// Mitsubishi GX Works2 project: V3 (working)   PLC: FX3U/FX3UC

PROGRAM MAIN
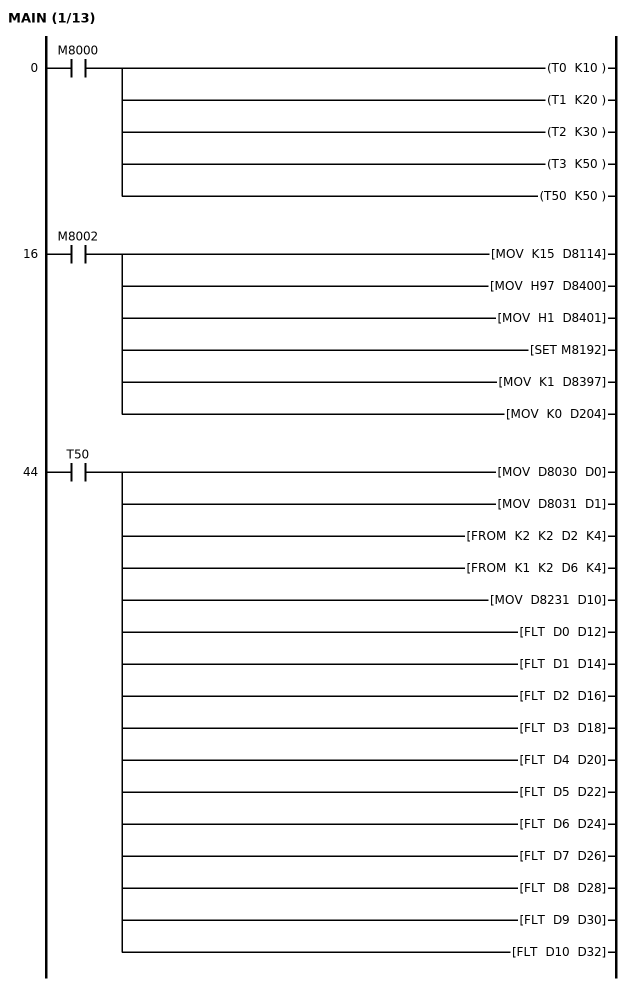
0     LD      M8000
      OUT     T0 K10
      OUT     T1 K20
      OUT     T2 K30
      OUT     T3 K50
      OUT     T50 K50
16    LD      M8002
      MOV     K15 D8114
      MOV     H97 D8400
      MOV     H1 D8401
      SET     M8192
      MOV     K1 D8397
      MOV     K0 D204
44    LD      T50
      MOV     D8030 D0
      MOV     D8031 D1
      FROM    K2 K2 D2 K4
      FROM    K1 K2 D6 K4
      MOV     D8231 D10
      FLT     D0 D12
      FLT     D1 D14
      FLT     D2 D16
      FLT     D3 D18
      FLT     D4 D20
      FLT     D5 D22
      FLT     D6 D24
      FLT     D7 D26
      FLT     D8 D28
      FLT     D9 D30
      FLT     D10 D32
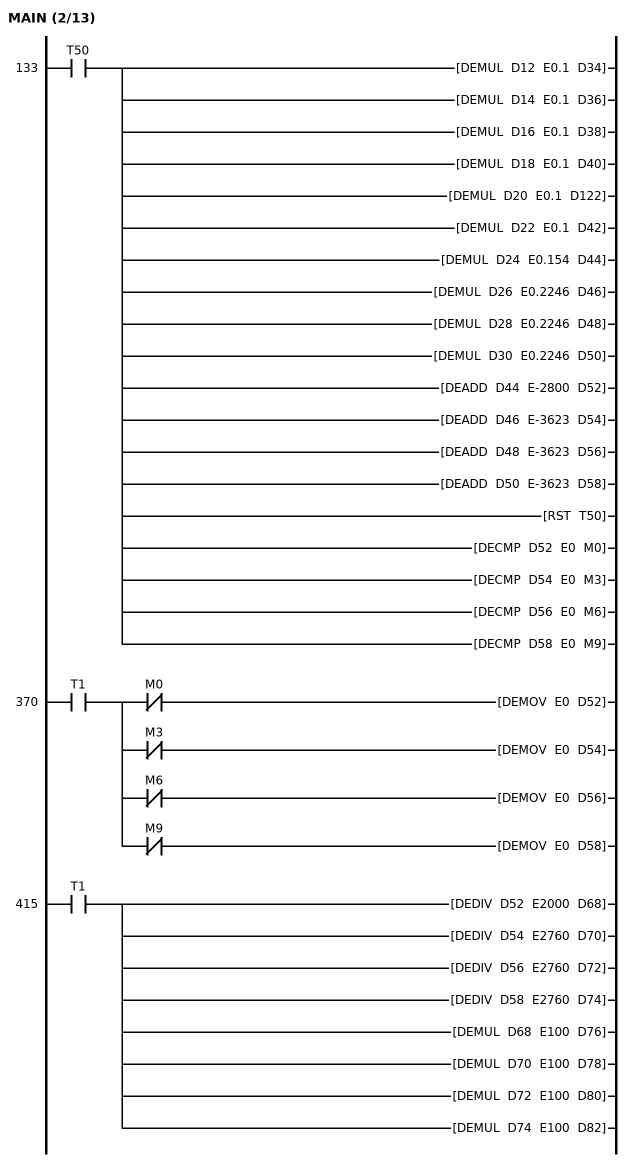
133   LD      T50
      DEMUL   D12 E0.1 D34
      DEMUL   D14 E0.1 D36
      DEMUL   D16 E0.1 D38
      DEMUL   D18 E0.1 D40
      DEMUL   D20 E0.1 D122
      DEMUL   D22 E0.1 D42
      DEMUL   D24 E0.154 D44
      DEMUL   D26 E0.2246 D46
      DEMUL   D28 E0.2246 D48
      DEMUL   D30 E0.2246 D50
      DEADD   D44 E-2800 D52
      DEADD   D46 E-3623 D54
      DEADD   D48 E-3623 D56
      DEADD   D50 E-3623 D58
      RST     T50
      DECMP   D52 E0 M0
      DECMP   D54 E0 M3
      DECMP   D56 E0 M6
      DECMP   D58 E0 M9
370   LD      T1
      MPS
      ANI     M0
      DEMOV   E0 D52
      MRD
      ANI     M3
      DEMOV   E0 D54
      MRD
      ANI     M6
      DEMOV   E0 D56
      MPP
      ANI     M9
      DEMOV   E0 D58
415   LD      T1
      DEDIV   D52 E2000 D68
      DEDIV   D54 E2760 D70
      DEDIV   D56 E2760 D72
      DEDIV   D58 E2760 D74
      DEMUL   D68 E100 D76
      DEMUL   D70 E100 D78
      DEMUL   D72 E100 D80
      DEMUL   D74 E100 D82
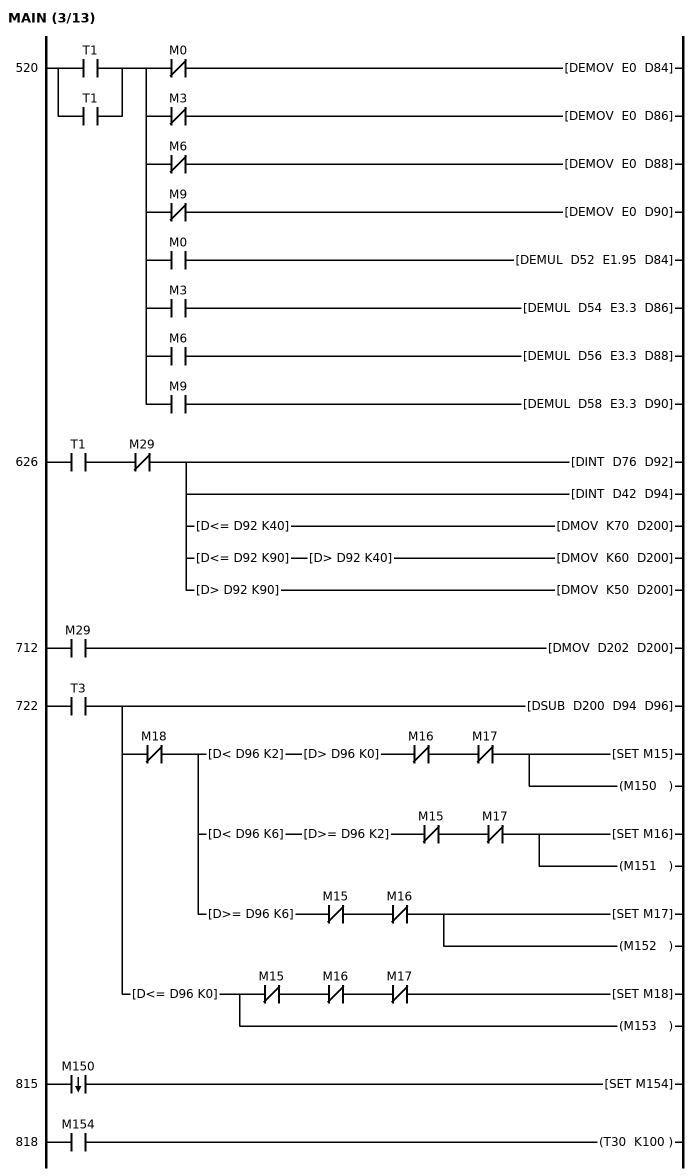
520   LD      T1
      OR      T1
      MPS
      ANI     M0
      DEMOV   E0 D84
      MRD
      ANI     M3
      DEMOV   E0 D86
      MRD
      ANI     M6
      DEMOV   E0 D88
      MRD
      ANI     M9
      DEMOV   E0 D90
      MRD
      AND     M0
      DEMUL   D52 E1.95 D84
      MRD
      AND     M3
      DEMUL   D54 E3.3 D86
      MRD
      AND     M6
      DEMUL   D56 E3.3 D88
      MPP
      AND     M9
      DEMUL   D58 E3.3 D90
626   LD      T1
      ANI     M29
      DINT    D76 D92
      DINT    D42 D94
      MPS
      ANDD<=  D92 K40
      DMOV    K70 D200
      MRD
      ANDD<=  D92 K90
      ANDD>   D92 K40
      DMOV    K60 D200
      MPP
      ANDD>   D92 K90
      DMOV    K50 D200
712   LD      M29
      DMOV    D202 D200
722   LD      T3
      DSUB    D200 D94 D96
      MPS
      ANI     M18
      MPS
      ANDD<   D96 K2
      ANDD>   D96 K0
      ANI     M16
      ANI     M17
      SET     M15
      OUT     M150
      MRD
      ANDD<   D96 K6
      ANDD>=  D96 K2
      ANI     M15
      ANI     M17
      SET     M16
      OUT     M151
      MPP
      ANDD>=  D96 K6
      ANI     M15
      ANI     M16
      SET     M17
      OUT     M152
      MPP
      ANDD<=  D96 K0
      MPS
      ANI     M15
      ANI     M16
      ANI     M17
      SET     M18
      MPP
      OUT     M153
815   LDF     M150
      SET     M154
818   LD      M154
      OUT     T30 K100
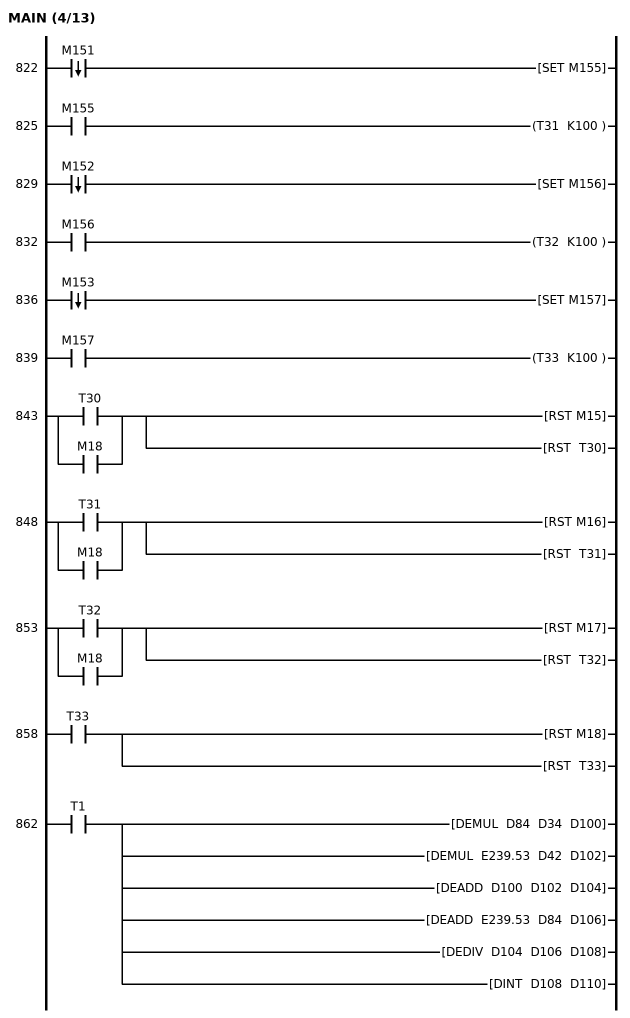
822   LDF     M151
      SET     M155
825   LD      M155
      OUT     T31 K100
829   LDF     M152
      SET     M156
832   LD      M156
      OUT     T32 K100
836   LDF     M153
      SET     M157
839   LD      M157
      OUT     T33 K100
843   LD      T30
      OR      M18
      RST     M15
      RST     T30
848   LD      T31
      OR      M18
      RST     M16
      RST     T31
853   LD      T32
      OR      M18
      RST     M17
      RST     T32
858   LD      T33
      RST     M18
      RST     T33
862   LD      T1
      DEMUL   D84 D34 D100
      DEMUL   E239.53 D42 D102
      DEADD   D100 D102 D104
      DEADD   E239.53 D84 D106
      DEDIV   D104 D106 D108
      DINT    D108 D110
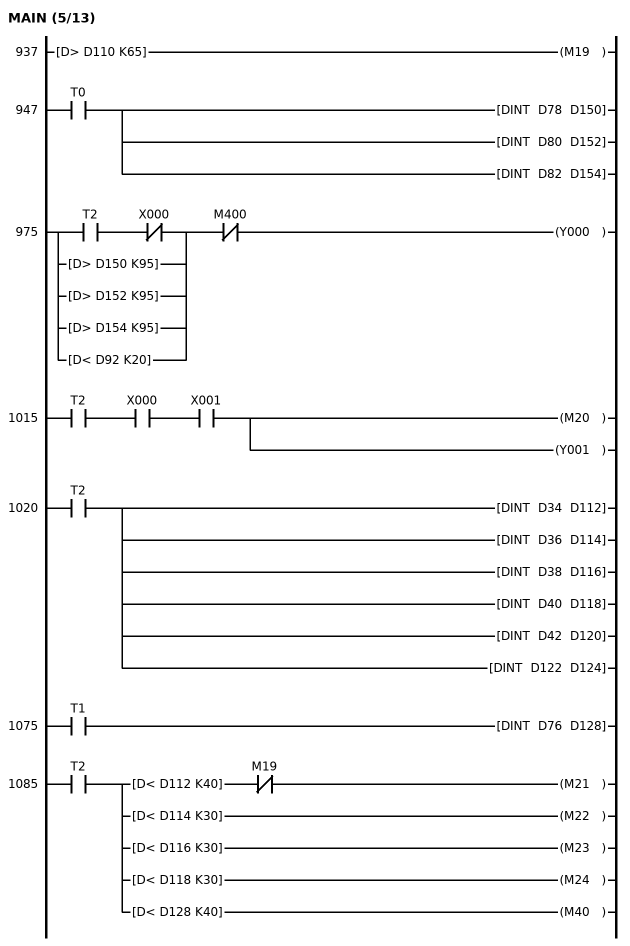
937   LDD>    D110 K65
      OUT     M19
947   LD      T0
      DINT    D78 D150
      DINT    D80 D152
      DINT    D82 D154
975   LD      T2
      ANI     X000
      ORD>    D150 K95
      ORD>    D152 K95
      ORD>    D154 K95
      ORD<    D92 K20
      ANI     M400
      OUT     Y000
1015  LD      T2
      AND     X000
      AND     X001
      OUT     M20
      OUT     Y001
1020  LD      T2
      DINT    D34 D112
      DINT    D36 D114
      DINT    D38 D116
      DINT    D40 D118
      DINT    D42 D120
      DINT    D122 D124
1075  LD      T1
      DINT    D76 D128
1085  LD      T2
      MPS
      ANDD<   D112 K40
      ANI     M19
      OUT     M21
      MRD
      ANDD<   D114 K30
      OUT     M22
      MRD
      ANDD<   D116 K30
      OUT     M23
      MRD
      ANDD<   D118 K30
      OUT     M24
      MPP
      ANDD<   D128 K40
      OUT     M40
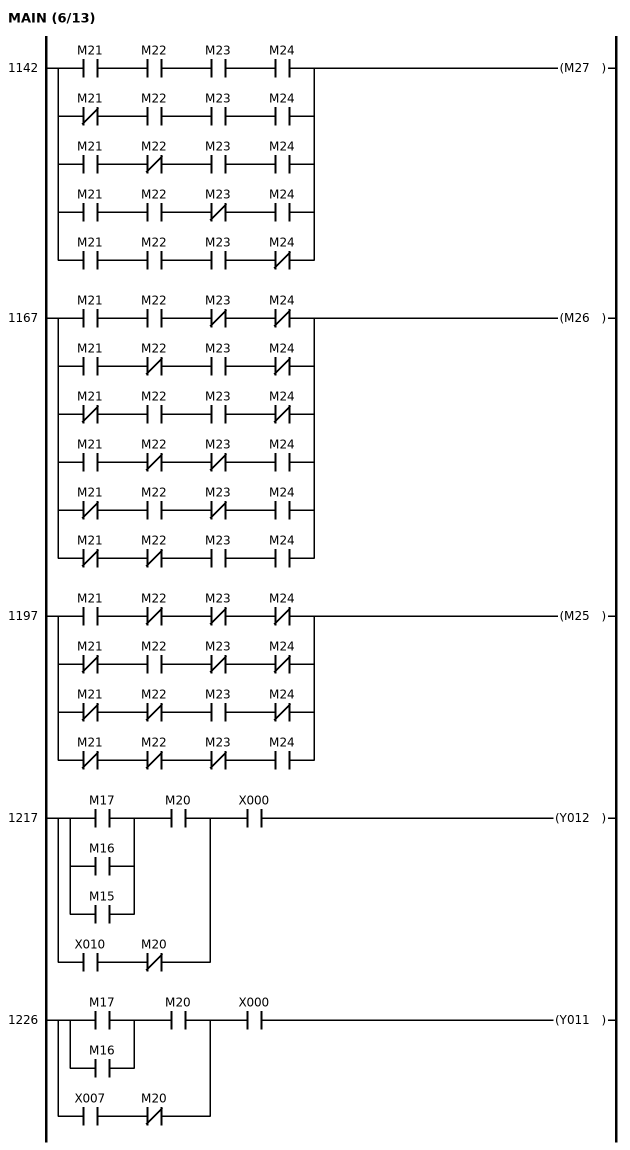
1142  LD      M21
      AND     M22
      AND     M23
      AND     M24
      LDI     M21
      AND     M22
      AND     M23
      AND     M24
      ORB
      LD      M21
      ANI     M22
      AND     M23
      AND     M24
      ORB
      LD      M21
      AND     M22
      ANI     M23
      AND     M24
      ORB
      LD      M21
      AND     M22
      AND     M23
      ANI     M24
      ORB
      OUT     M27
1167  LD      M21
      AND     M22
      ANI     M23
      ANI     M24
      LD      M21
      ANI     M22
      AND     M23
      ANI     M24
      ORB
      LDI     M21
      AND     M22
      AND     M23
      ANI     M24
      ORB
      LD      M21
      ANI     M22
      ANI     M23
      AND     M24
      ORB
      LDI     M21
      AND     M22
      ANI     M23
      AND     M24
      ORB
      LDI     M21
      ANI     M22
      AND     M23
      AND     M24
      ORB
      OUT     M26
1197  LD      M21
      ANI     M22
      ANI     M23
      ANI     M24
      LDI     M21
      AND     M22
      ANI     M23
      ANI     M24
      ORB
      LDI     M21
      ANI     M22
      AND     M23
      ANI     M24
      ORB
      LDI     M21
      ANI     M22
      ANI     M23
      AND     M24
      ORB
      OUT     M25
1217  LD      M17
      OR      M16
      OR      M15
      AND     M20
      LD      X010
      ANI     M20
      ORB
      AND     X000
      OUT     Y012
1226  LD      M17
      OR      M16
      AND     M20
      LD      X007
      ANI     M20
      ORB
      AND     X000
      OUT     Y011
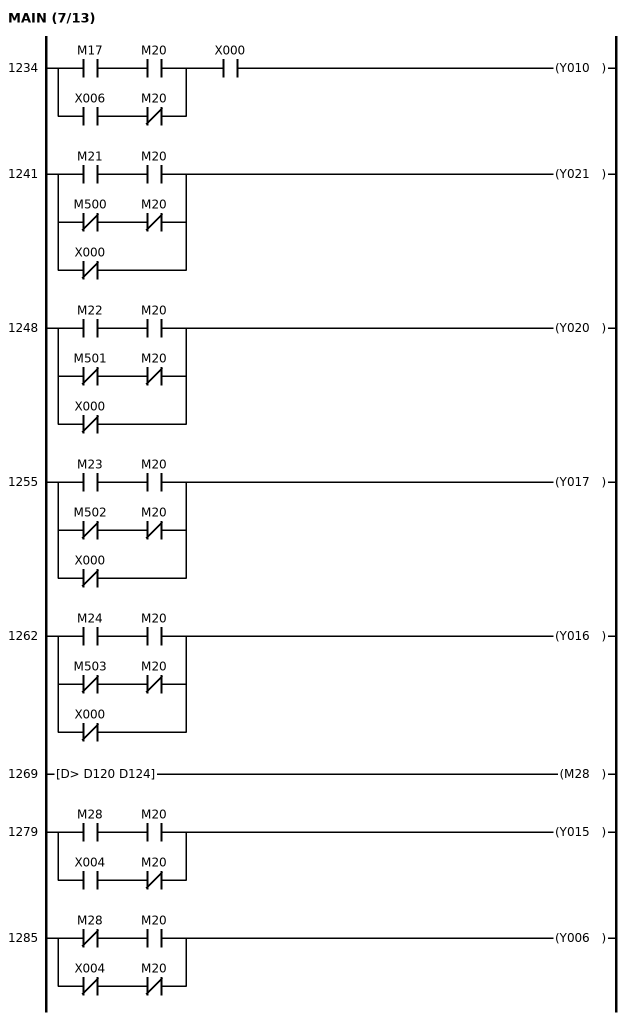
1234  LD      M17
      AND     M20
      LD      X006
      ANI     M20
      ORB
      AND     X000
      OUT     Y010
1241  LD      M21
      AND     M20
      LDI     M500
      ANI     M20
      ORB
      ORI     X000
      OUT     Y021
1248  LD      M22
      AND     M20
      LDI     M501
      ANI     M20
      ORB
      ORI     X000
      OUT     Y020
1255  LD      M23
      AND     M20
      LDI     M502
      ANI     M20
      ORB
      ORI     X000
      OUT     Y017
1262  LD      M24
      AND     M20
      LDI     M503
      ANI     M20
      ORB
      ORI     X000
      OUT     Y016
1269  LDD>    D120 D124
      OUT     M28
1279  LD      M28
      AND     M20
      LD      X004
      ANI     M20
      ORB
      OUT     Y015
1285  LDI     M28
      AND     M20
      LDI     X004
      ANI     M20
      ORB
      OUT     Y006
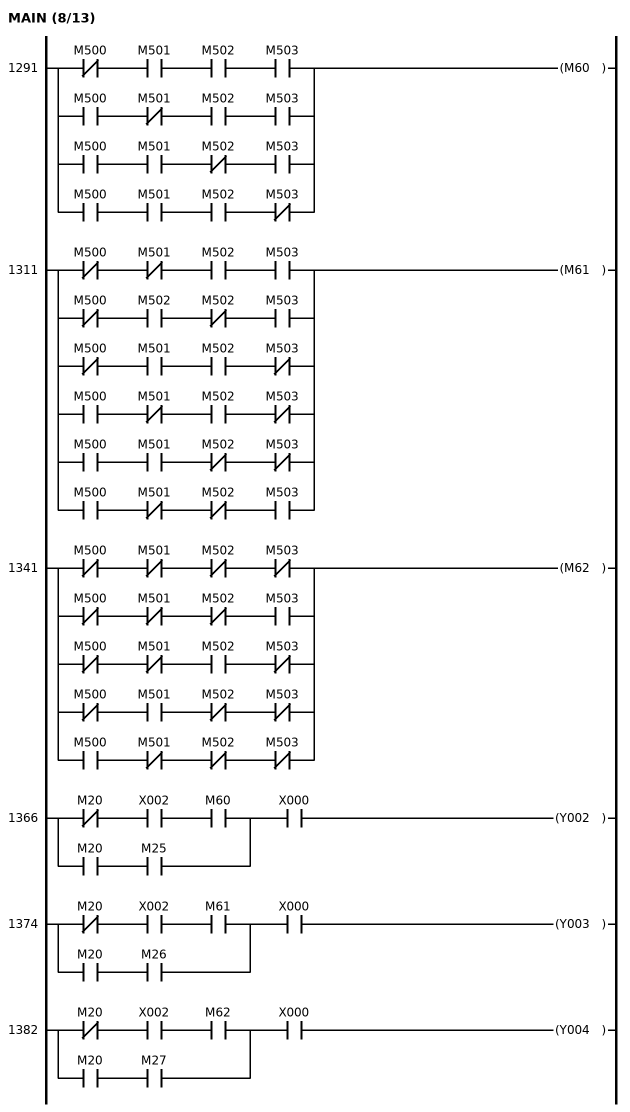
1291  LDI     M500
      AND     M501
      AND     M502
      AND     M503
      LD      M500
      ANI     M501
      AND     M502
      AND     M503
      ORB
      LD      M500
      AND     M501
      ANI     M502
      AND     M503
      ORB
      LD      M500
      AND     M501
      AND     M502
      ANI     M503
      ORB
      OUT     M60
1311  LDI     M500
      ANI     M501
      AND     M502
      AND     M503
      LDI     M500
      AND     M502
      ANI     M502
      AND     M503
      ORB
      LDI     M500
      AND     M501
      AND     M502
      ANI     M503
      ORB
      LD      M500
      ANI     M501
      AND     M502
      ANI     M503
      ORB
      LD      M500
      AND     M501
      ANI     M502
      ANI     M503
      ORB
      LD      M500
      ANI     M501
      ANI     M502
      AND     M503
      ORB
      OUT     M61
1341  LDI     M500
      ANI     M501
      ANI     M502
      ANI     M503
      LDI     M500
      ANI     M501
      ANI     M502
      AND     M503
      ORB
      LDI     M500
      ANI     M501
      AND     M502
      ANI     M503
      ORB
      LDI     M500
      AND     M501
      ANI     M502
      ANI     M503
      ORB
      LD      M500
      ANI     M501
      ANI     M502
      ANI     M503
      ORB
      OUT     M62
1366  LDI     M20
      AND     X002
      AND     M60
      LD      M20
      AND     M25
      ORB
      AND     X000
      OUT     Y002
1374  LDI     M20
      AND     X002
      AND     M61
      LD      M20
      AND     M26
      ORB
      AND     X000
      OUT     Y003
1382  LDI     M20
      AND     X002
      AND     M62
      LD      M20
      AND     M27
      ORB
      AND     X000
      OUT     Y004
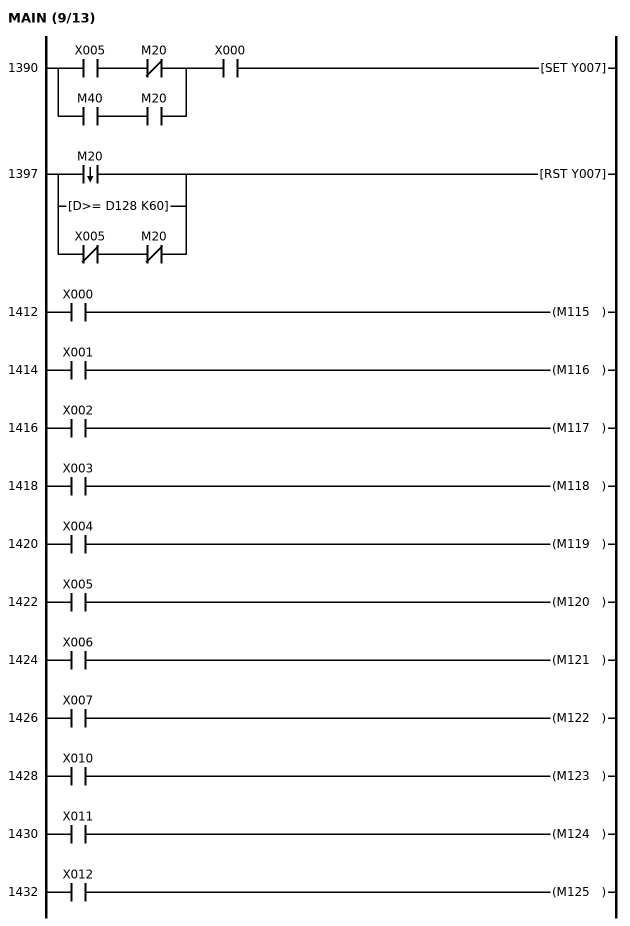
1390  LD      X005
      ANI     M20
      LD      M40
      AND     M20
      ORB
      AND     X000
      SET     Y007
1397  LDF     M20
      ORD>=   D128 K60
      LDI     X005
      ANI     M20
      ORB
      RST     Y007
1412  LD      X000
      OUT     M115
1414  LD      X001
      OUT     M116
1416  LD      X002
      OUT     M117
1418  LD      X003
      OUT     M118
1420  LD      X004
      OUT     M119
1422  LD      X005
      OUT     M120
1424  LD      X006
      OUT     M121
1426  LD      X007
      OUT     M122
1428  LD      X010
      OUT     M123
1430  LD      X011
      OUT     M124
1432  LD      X012
      OUT     M125
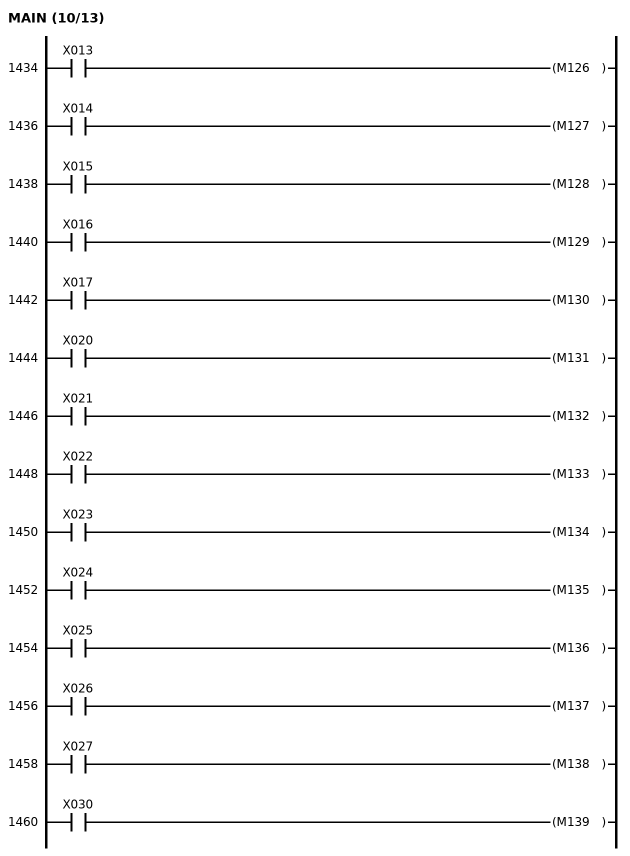
1434  LD      X013
      OUT     M126
1436  LD      X014
      OUT     M127
1438  LD      X015
      OUT     M128
1440  LD      X016
      OUT     M129
1442  LD      X017
      OUT     M130
1444  LD      X020
      OUT     M131
1446  LD      X021
      OUT     M132
1448  LD      X022
      OUT     M133
1450  LD      X023
      OUT     M134
1452  LD      X024
      OUT     M135
1454  LD      X025
      OUT     M136
1456  LD      X026
      OUT     M137
1458  LD      X027
      OUT     M138
1460  LD      X030
      OUT     M139
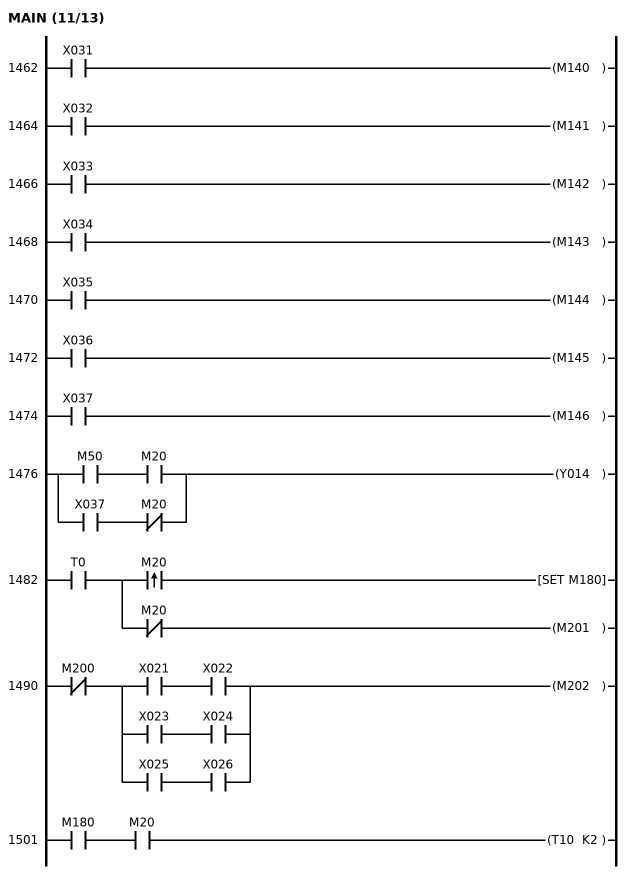
1462  LD      X031
      OUT     M140
1464  LD      X032
      OUT     M141
1466  LD      X033
      OUT     M142
1468  LD      X034
      OUT     M143
1470  LD      X035
      OUT     M144
1472  LD      X036
      OUT     M145
1474  LD      X037
      OUT     M146
1476  LD      M50
      AND     M20
      LD      X037
      ANI     M20
      ORB
      OUT     Y014
1482  LD      T0
      MPS
      ANDP    M20
      SET     M180
      MPP
      ANI     M20
      OUT     M201
1490  LDI     M200
      LD      X021
      AND     X022
      LD      X023
      AND     X024
      ORB
      LD      X025
      AND     X026
      ORB
      ANB
      OUT     M202
1501  LD      M180
      AND     M20
      OUT     T10 K2
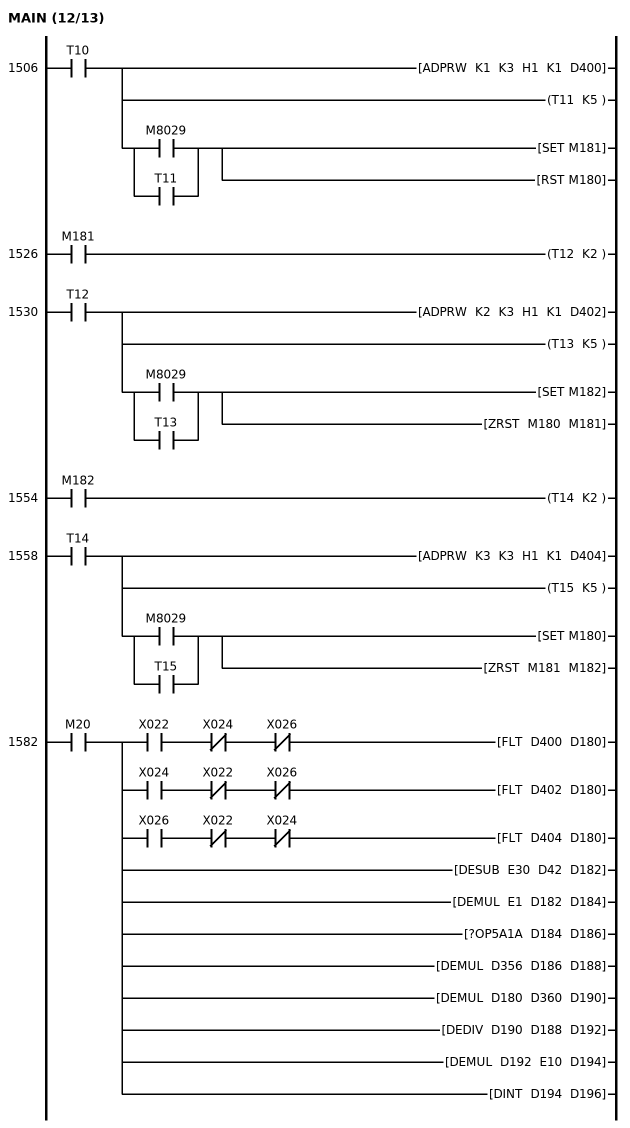
1506  LD      T10
      ADPRW   K1 K3 H1 K1 D400
      OUT     T11 K5
      LD      M8029
      OR      T11
      ANB
      SET     M181
      RST     M180
1526  LD      M181
      OUT     T12 K2
1530  LD      T12
      ADPRW   K2 K3 H1 K1 D402
      OUT     T13 K5
      LD      M8029
      OR      T13
      ANB
      SET     M182
      ZRST    M180 M181
1554  LD      M182
      OUT     T14 K2
1558  LD      T14
      ADPRW   K3 K3 H1 K1 D404
      OUT     T15 K5
      LD      M8029
      OR      T15
      ANB
      SET     M180
      ZRST    M181 M182
1582  LD      M20
      MPS
      AND     X022
      ANI     X024
      ANI     X026
      FLT     D400 D180
      MRD
      AND     X024
      ANI     X022
      ANI     X026
      FLT     D402 D180
      MRD
      AND     X026
      ANI     X022
      ANI     X024
      FLT     D404 D180
      MPP
      DESUB   E30 D42 D182
      DEMUL   E1 D182 D184
      ?OP5A1A D184 D186
      DEMUL   D356 D186 D188
      DEMUL   D180 D360 D190
      DEDIV   D190 D188 D192
      DEMUL   D192 E10 D194
      DINT    D194 D196
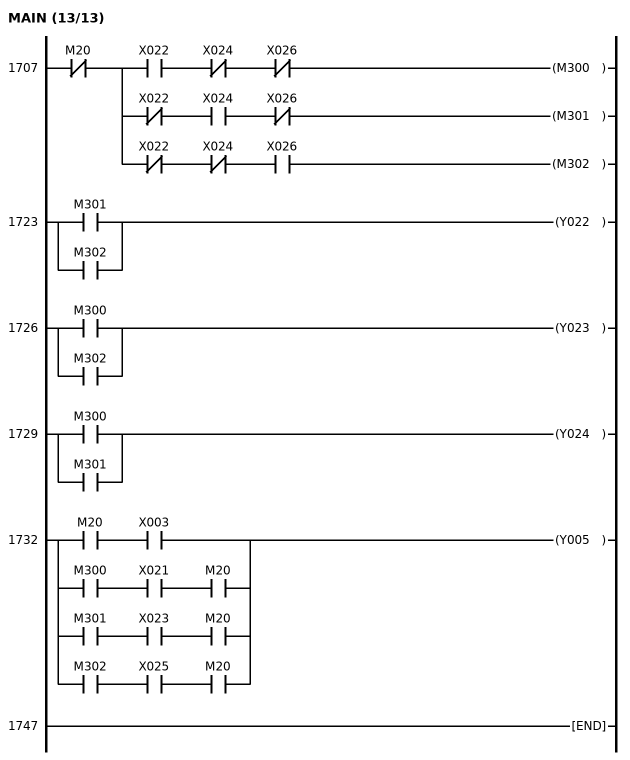
1707  LDI     M20
      MPS
      AND     X022
      ANI     X024
      ANI     X026
      OUT     M300
      MRD
      ANI     X022
      AND     X024
      ANI     X026
      OUT     M301
      MPP
      ANI     X022
      ANI     X024
      AND     X026
      OUT     M302
1723  LD      M301
      OR      M302
      OUT     Y022
1726  LD      M300
      OR      M302
      OUT     Y023
1729  LD      M300
      OR      M301
      OUT     Y024
1732  LD      M20
      AND     X003
      LD      M300
      AND     X021
      AND     M20
      ORB
      LD      M301
      AND     X023
      AND     M20
      ORB
      LD      M302
      AND     X025
      AND     M20
      ORB
      OUT     Y005
1747  END
END_PROGRAM
